Staubli VAL3: savePROG.dtx

public progItem pProgItem{}
  [Key1]
    progTemplate pProgTemplate
      [0]
        string sTRAJname
        num nType
        ifItem iIfItem
          [0]
            num nSigType[3]
            num nSigIndex[3]
            num nValue[3]
            bool bANDOR[2]
        switchItem sSwitchItem
          [0]
            num nSwitchValue
            string sIOValue
            bool bIOdisable
        forItem fForItem
          [0]
            num nLoopValue
            bool bIOdisable
            string sIOindex
